// TIA Portal V20 export
Screen "Pop-up_SafetyGate"  395x590
  ScreenItem "Text field TG Status" at 1,0 size 394x47  Type=HmiTextBox
  ScreenItem "Cancel Mode" at 315,3 size 76x42  Type=HmiButton
  ScreenItem "Background_1" at 0,37 size 368x32  Type=HmiRectangle
  ScreenItem "Text field TG1 Status_22" at 51,43 size 126x21  Type=HmiTextBox
  ScreenItem "Text field TG1 Status_1" at 191,43 size 78x21  Type=HmiTextBox
  ScreenItem "Rectangle TG1" at 1,74 size 367x40  Type=HmiRectangle
  ScreenItem "Textfeld_1" at 7,83 size 140x20  Type=HmiTextBox
  ScreenItem "Textfeld_2" at 155,83 size 245x20  Type=HmiTextBox
  ScreenItem "Rectangle TG1_1" at 1,115 size 367x40  Type=HmiRectangle
  ScreenItem "Rectangle TG1_2" at 1,156 size 367x40  Type=HmiRectangle
  ScreenItem "Rectangle TG1_3" at 1,238 size 367x40  Type=HmiRectangle
  ScreenItem "Rectangle TG1_4" at 1,197 size 367x40  Type=HmiRectangle
  ScreenItem "Textfeld_10" at 7,121 size 140x20  Type=HmiTextBox
  ScreenItem "Textfeld_13" at 155,121 size 275x20  Type=HmiTextBox
  ScreenItem "Textfeld_5" at 7,161 size 140x20  Type=HmiTextBox
  ScreenItem "Textfeld_14" at 156,161 size 275x20  Type=HmiTextBox
  ScreenItem "Textfeld_6" at 7,206 size 140x20  Type=HmiTextBox
  ScreenItem "Textfeld_15" at 161,206 size 110x20  Type=HmiTextBox
  ScreenItem "Textfeld_8" at 7,249 size 140x20  Type=HmiTextBox
  ScreenItem "Textfeld_21" at 155,249 size 275x20  Type=HmiTextBox
  ScreenItem "Line_1" at 152,74 size 1x203  Type=HmiLine
  ScreenItem "Background_2" at 0,0 size 368x32  Type=HmiRectangle
  ScreenItem "Text field TG1 Status_2" at 142,7 size 126x21  Type=HmiTextBox
  ScreenItem "Background_3" at 12,382 size 368x32  Type=HmiRectangle
  ScreenItem "Text field TG1 Status_4" at 63,388 size 126x21  Type=HmiTextBox
  ScreenItem "Text field TG1 Status_3" at 203,388 size 78x21  Type=HmiTextBox
  ScreenItem "Rectangle TG1_8" at 13,419 size 367x40  Type=HmiRectangle
  ScreenItem "Textfeld_19" at 19,428 size 140x20  Type=HmiTextBox
  ScreenItem "Textfeld_18" at 167,428 size 245x20  Type=HmiTextBox
  ScreenItem "Rectangle TG1_7" at 13,460 size 367x40  Type=HmiRectangle
  ScreenItem "Rectangle TG1_6" at 13,501 size 367x40  Type=HmiRectangle
  ScreenItem "Rectangle TG1_9" at 13,542 size 367x40  Type=HmiRectangle
  ScreenItem "Textfeld_16" at 167,466 size 275x20  Type=HmiTextBox
  ScreenItem "Textfeld_12" at 19,506 size 140x20  Type=HmiTextBox
  ScreenItem "Textfeld_11" at 168,506 size 275x20  Type=HmiTextBox
  ScreenItem "Textfeld_9" at 19,551 size 140x20  Type=HmiTextBox
  ScreenItem "Textfeld_7" at 173,551 size 133x20  Type=HmiTextBox
  ScreenItem "Line_2" at 164,419 size 2x163  Type=HmiLine
  ScreenItem "Background_4" at 12,345 size 368x32  Type=HmiRectangle
  ScreenItem "Text field TG1 Status_5" at 109,352 size 197x21  Type=HmiTextBox
  ScreenItem "Textfeld_3" at 20,468 size 140x20  Type=HmiTextBox
